// TIA Portal V19 export
// export: Created 2026-11-08T08:30:00.0000000Z, ExportSetting WithReadOnly, DisplayName Totally Integrated Automation Portal, DisplayVersion V19
FUNCTION_BLOCK "FB_ExampleValve"   // FB10, SCL
{ S7_Optimized_Access := 'TRUE' }
VERSION : 0.1
// Example valve block (synthetic)
// stored: AutoNumber true, CodeModifiedDate 2026-01-10T09:00:00.0000000Z, CompileDate 2026-01-10T09:05:00.0000000Z, IsConsistent true, IsIECCheckEnabled false, IsKnowHowProtected false, ModifiedDate 2026-01-10T09:00:00.0000000Z, SetENOAutomatically false
   VAR_INPUT
      Open : Bool;   // Open command
      Interlock : Bool;
   END_VAR
   VAR_OUTPUT
      Output : Bool;
   END_VAR
   VAR RETAIN
      OpenCount : DInt := 0;
   END_VAR
   VAR
      Limit : Real := 90.0;
   END_VAR
   VAR CONSTANT
      MaxCount : DInt := 1000;
   END_VAR
BEGIN
// Valve logic
   // Example valve permissive
   IF #Open AND NOT #Interlock THEN
       #Output := TRUE;
       #OpenCount := #OpenCount + 1; (*count openings*)
   ELSE
       #Output := FALSE;
   END_IF;
END_FUNCTION_BLOCK
